Fanuc KAREL source: KT00533.KL

PROGRAM KT00533
%NOLOCKGROUP
VAR
  P1: JOINTPOS
  P2: POSITION
  OUT: BOOLEAN
BEGIN
  OUT = P1 >=< P2
END KT00533
